Staubli VAL3: switchItem.dtx

public num nSwitchValue
public string sIOValue
public bool bIOdisable
